Universal Robots PolyScope program: PrecProg.urp

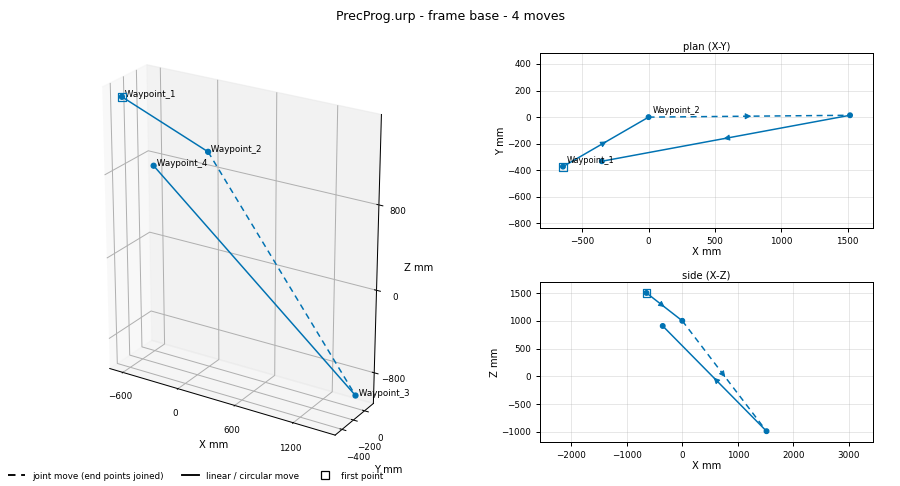
[picture p0: tool path of PrecProg.urp in frame base, 4 of 4 moves have a stored position in this frame; points joined in program order, loops and branches not executed]
Program PrecProg (createdIn=3.0.0 lastSavedIn=3.0.0 directory=/programs installation=default)
Robot Program (runOnlyOnce=true motionType=MoveJ speed=1.047198 acceleration=1.396263 useActiveTCP=false)
  'Program generated by RoboDK v6.0.7 for ABB IRB 120-3/0.6 on XX/XX/XXXX 18:00:00'
  'Using nominal kinematics.'
  'Using Ref. Frame P: p[0.000000, -0.000001, 1.000000, 1.570792, -0.005162, 0.008546]'
  'Using TCP Tool P: p[0.000125, -0.000375, 0.123457, -0.789761, -0.000001, 0.000002]'
  Script: set_tcp(p[0.000125, -0.000375, 0.123457, -0.789761, -0.000001, 0.000002])
  Script: movej([0.215471, -0.797247, 1.377087, -0.008727, 0.008726, 3.141593],1.20000,0.75000,0,0.0000)
  MoveL speed 250 mm/s, acceleration 1200 mm/s^2 (useActiveTCP=true)
    Waypoint Waypoint_1: TCP in base x=-644.182 y=-372.923 z=1501.372 mm, rx=1.3972 ry=2.2886 rz=1.3609 rad; joints [12.346, -45.679, 78.901, -0.5, 0.5, 180] deg; flange x=-632.669 y=-412.763 z=1617.656 mm, rx=-1.3289 ry=-2.5613 rz=-0.3651 rad
    Waypoint Waypoint_2: TCP in base x=0.505 y=-0.25 z=999.504 mm, rx=-1.5708 ry=-0.0085 rz=-0.0053 rad; joints [-12.345, 45.678, -78.9, 0.5, 0, -180] deg; flange x=1.334 y=-86.897 z=911.565 mm, rx=-0.781 ry=-0.0092 rz=-0.0015 rad
  Script: movej([-0.215468, 0.797240, -1.377065, 0.008727, -0.000002, -3.141593],1.20000,0.75000,0,0.0000)
  MoveJ speed 42.97 deg/s, acceleration 68.75 deg/s^2 (useActiveTCP=true)
    Waypoint Waypoint_3: TCP in base x=1517.499 y=13.766 z=-987.823 mm, rx=1.2018 ry=1.2044 rz=1.2149 rad; joints [-12.345, 45.678, -78.9, 0.5, 0, -180] deg; flange x=1430.086 y=13.452 z=-900.641 mm, rx=1.7555 ry=1.7593 rz=0.7332 rad
  Script: movej([-0.215468, 0.797240, -1.377065, 0.008727, -0.000002, -3.141593],1.20000,0.75000,0,0.0000)
  Wait Sleep waitTime=0.002
  Wait Sleep waitTime=1
  MoveL speed 67 mm/s, acceleration 1200 mm/s^2 (useActiveTCP=true)
    Waypoint Waypoint_4: TCP in base x=-351.51 y=-332.461 z=906.789 mm, rx=0.7612 ry=2.0119 rz=1.6554 rad; joints [12.346, -45.679, 78.901, -0.5, 0.5, 180] deg; flange x=-393.645 y=-385.039 z=1010.239 mm, rx=0.9946 ry=2.6694 rz=0.8071 rad
